{attribute 'qualified_only'}
VAR_GLOBAL PERSISTENT
    sMqttPassword : STRING(63);                                  // empty = telemetry stays offline
    aEnergyWh     : ARRAY[1..GVL_Param.FEED_COUNT] OF LREAL;     // Wh per feed since local midnight
    nEnergyDay    : UDINT;                                       // local day number the counters belong to
END_VAR

(* stored: Version 1.1.0.1
   GVL GVL_Persist: Id {37ce5e80-ae4b-490d-b27a-ae2eb12b868e} *)
